TEXTLIST TextList_CIP_Clients
  0 = ' '
  1 = 'Tank1 Marinada'
  2 = 'Tank2 Marinada'
  3 = 'Tank3 Color'
  4 = 'Tank4 Color'
  5 = 'TriBlender Marinada'
  6 = 'TriBlender Color'
  7 = 'Line Marinada'
  8 = 'Line Color'
  9 = 'Local'
   = ''
END_TEXTLIST

(* stored: Version 1.1.0.1, ProductVersion 3.1.4024.12
   TextList TextList_CIP_Clients: Id {efff2837-8fe3-4cf4-ac8f-92f682fb3c49} *)
